(* IEC 61131-3 sources: plc-st-coding-agent/progress/evidence/review_r8_first_candidate_20261110_v2/native_artifacts/codex_deepseek-v4pro/self-medium-03, 1 file *)

(* ---- candidate.st ---- *)
FUNCTION_BLOCK FB
VAR_INPUT
    openBtn: BOOL;
    closeBtn: BOOL;
    openLimit: BOOL;
    closeLimit: BOOL;
    obstacle: BOOL;
END_VAR
VAR_OUTPUT
    motorUp: BOOL;
    motorDown: BOOL;
    errorFlag: BOOL;
END_VAR
VAR
    prevOpenBtn: BOOL;
    prevCloseBtn: BOOL;
    prevMotorUp: BOOL;
    prevMotorDown: BOOL;
    prevErrorFlag: BOOL;
    openRising: BOOL;
    closeRising: BOOL;
    bothRising: BOOL;
END_VAR

openRising := openBtn AND NOT prevOpenBtn;
closeRising := closeBtn AND NOT prevCloseBtn;
bothRising := openBtn AND closeBtn AND NOT (prevOpenBtn AND prevCloseBtn);

errorFlag := obstacle OR (prevErrorFlag AND NOT bothRising);

motorUp := NOT obstacle AND NOT openLimit AND
           (prevMotorUp OR
            (NOT prevMotorUp AND NOT prevMotorDown AND NOT prevErrorFlag AND openRising AND NOT closeBtn));

motorDown := NOT obstacle AND NOT closeLimit AND
             (prevMotorDown OR
              (NOT prevMotorUp AND NOT prevMotorDown AND NOT prevErrorFlag AND closeRising AND NOT openBtn));

prevOpenBtn := openBtn;
prevCloseBtn := closeBtn;
prevMotorUp := motorUp;
prevMotorDown := motorDown;
prevErrorFlag := errorFlag;
END_FUNCTION_BLOCK
